// TIA Portal V20 export
TYPE "Kistler_Fertigungsauftragsnummer"
   STRUCT
      Fertigungauftragsnummer : Array[0..25] of Char;
   END_STRUCT;
END_TYPE
